Fanuc KAREL source: KO00028.KL

PROGRAM KO00028
%NOLOCKGROUP
VAR
  P1: JOINTPOS
  P2: JOINTPOS
  P3: JOINTPOS
  OUT: JOINTPOS
BEGIN
  OUT = FRAME(P1, P2, P3)
END KO00028
